FUNCTION_BLOCK ConveyorPointHMI (* CAT Function Block Type *)
  (* Standard: 61499-2 *)
  (* Version 0.0, 7/9/2026, template *)
  PACKAGE Main;
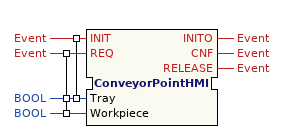
  EVENT_INPUT
    INIT WITH Tray; (* Initialization Request *)
    REQ WITH Tray, Workpiece; (* Normal Execution Request *)
  END_EVENT
  EVENT_OUTPUT
    INITO; (* Initialization Confirm *)
    CNF; (* Execution Confirmation *)
    RELEASE;
  END_EVENT
  VAR_INPUT
    Tray : BOOL; (* Input event qualifier *)
    Workpiece : BOOL;
  END_VAR
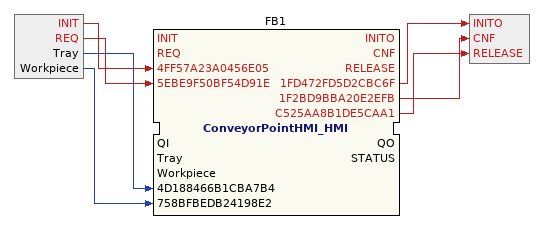
  FBS
    FB1 : ConveyorPointHMI_HMI;
  END_FBS
  EVENT_CONNECTIONS
    INIT TO FB1.4FF57A23A0456E05;
    REQ TO FB1.5EBE9F50BF54D91E;
    FB1.1FD472FD5D2CBC6F TO INITO;
    FB1.1F2BD9BBA20E2EFB TO CNF;
    FB1.C525AA8B1DE5CAA1 TO RELEASE;
  END_CONNECTIONS
  DATA_CONNECTIONS
    Tray TO FB1.4D188466B1CBA7B4;
    Workpiece TO FB1.758BFBEDB24198E2;
  END_CONNECTIONS
END_FUNCTION_BLOCK
